// TIA Portal V21 export
// export: Created 2026-10-08T11:46:22.7242637Z, ExportSetting WithDefaults, DisplayName Totally Integrated Automation Portal, DisplayVersion V21 Update 2, DisplayName TIA Portal Test Suite Advanced, DisplayVersion V21, DisplayName SINAMICS Startdrive Advanced, DisplayVersion V21 HF2, DisplayName SINAMICS DCC, DisplayVersion V21, DisplayName SINAMICS Startdrive G110M, G120, G120C, G120D, G120P, G115D, DisplayVersion V21 HF2, DisplayName SINAMICS Startdrive G130, G150, S120, S150, G200, G220, S200, S210, S220, Innomotics MVD, DisplayVersion V21 HF2, DisplayName STEP 7 Professional, DisplayVersion V21 Update 2, DisplayName STEP 7 Safety, DisplayVersion V21, DisplayName Tech WebApplication, DisplayVersion V21, DisplayName WinCC Basic/Comfort/Advanced, DisplayVersion V21 Update 2, DisplayName WinCC Unified, DisplayVersion V21 Update 2
FUNCTION_BLOCK "TgpUnit_TP_FBD"   // FB616, FBD
VERSION : 0.1
// stored: Access Unpublished, AutoNumber true, IsIECCheckEnabled false, IsRetainMemResEnabled false, MemoryReserve 100, Namespace TiaMcp_UnitA, SetENOAutomatically false, UDAEnableTagReadback false
   VAR_INPUT
      Enable : Bool;
      Preset : Time;
   END_VAR
   VAR_OUTPUT
      Done : Bool;
      Elapsed : Time;
   END_VAR
   VAR
      Storage { S7_SetPoint := 'True'} : TP_TIME;
   END_VAR
BEGIN

REGION Network 1
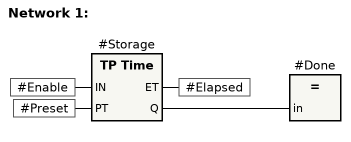
   #Storage(IN := #Enable, PT := #Preset, ET => #Elapsed);   // TP
   #Done := #Storage.Q;
END_REGION
END_FUNCTION_BLOCK
